Fanuc KAREL source: kt00136.KL

-- PROVISIONAL review KL for V940-1; original PC SHA256 3f5dac75cd2b1368fc149c27554bcc0b740e1e46f4c48efd419d121eed9d6ebe
-- Incomplete behavior may be omitted. Consult companion uncertainty JSON. Do not deploy.
PROGRAM KT00136
%NOLOCKGROUP
VAR
  I1 : INTEGER
  OUT : REAL
-- UNRESOLVED_DECL H2 type=002017
BEGIN
  -- V9_ZERO_TABLE_METADATA_HINT layout=0001; no indexed target words; source/name/runtime held
  -- UNRESOLVED_PC offsets 5-16; opcodes 2E,23
  -- UNRESOLVED_PC offsets 21-35; opcodes 2E,22,9D,33,B4
  -- UNRESOLVED_PC offsets 40-63; opcodes 21,22,9D,33,B3,55,64,23
  -- UNRESOLVED_PC offsets 68-72; opcodes 7F
END KT00136
